(* IEC 61131-3 sources: plc-process-lib/tests/POUs/Suites/FB_Motor_Test, 58 files *)

(* ---- AutoRunStartsAndConfirms.method.decl.st ---- *)
// Auto: запрос xAutoRun запускает двигатель (Starting, xQRun), ОС через 1 с подтверждает пуск (Running);
// пуск считается по фронту ОС, отметка в окне пусков — при входе в Starting; двигатель доступен автоматике.
METHOD PRIVATE AutoRunStartsAndConfirms
VAR
    fbTime   : FB_FakeTime;       // подменное время, старт 1 ч
    fbMot    : FB_Motor;          // двигатель под тестом
    stCmd    : ST_MotorCmd;       // команды
    stRetain : ST_DeviceRetain;   // энергонезависимые данные
    stCfg    : ST_MotorCfg;       // конфигурация (умолчания)
END_VAR

(* ---- CfgChecksSetEachCfgErrBit.method.decl.st ---- *)
// CheckConfig двигателя: каждая проверка 13.9 даёт свой бит wCfgErr; границы допустимы (30 пусков в час,
// tResetPulse = tResetWindow); без ОС времена ОС не проверяются.
METHOD PRIVATE CfgChecksSetEachCfgErrBit
VAR
    fbTime   : FB_FakeTime;       // подменное время, старт 1 ч
    fbMot    : FB_Motor;          // двигатель под тестом
    stCmd    : ST_MotorCmd;       // команды
    stRetain : ST_DeviceRetain;   // энергонезависимые данные
    stCfg    : ST_MotorCfg;       // конфигурация (умолчания)
    uBad     : U_TestEnumInt;     // значение вне перечисления
END_VAR

(* ---- CurrentRunSecondsCountsAndResetsOnStop.method.decl.st ---- *)
// Текущая непрерывная работа: 65 с работы — CurrentRunSeconds = 65 (и stSts.udiRunCurrent_s); останов — 0;
// новый пуск считает с нуля (3 с), наработка всего продолжается (68 с).
// Источник: tools/reference/motor.py, сценарии current_run_*.
METHOD PRIVATE CurrentRunSecondsCountsAndResetsOnStop
VAR
    fbTime   : FB_FakeTime;       // подменное время, старт 1 ч
    fbMot    : FB_Motor;          // двигатель под тестом
    stCmd    : ST_MotorCmd;       // команды
    stRetain : ST_DeviceRetain;   // энергонезависимые данные
    stCfg    : ST_MotorCfg;       // конфигурация (умолчания)
END_VAR

(* ---- ExtFaultInLocalLatches.method.decl.st ---- *)
// Внешняя авария действует и в Local: отказ фиксируется (Fault); после возврата в Manual отказ остаётся,
// пуск — RejectedFault.
METHOD PRIVATE ExtFaultInLocalLatches
VAR
    fbTime   : FB_FakeTime;       // подменное время, старт 1 ч
    fbMot    : FB_Motor;          // двигатель под тестом
    stCmd    : ST_MotorCmd;       // команды
    stRetain : ST_DeviceRetain;   // энергонезависимые данные
    stCfg    : ST_MotorCfg;       // конфигурация (умолчания)
END_VAR

(* ---- ExtFaultTripsAndResetRejectedWhileActive.method.decl.st ---- *)
// Внешняя авария через фильтр tExtFaultFilter = 200 мс: отказ ExtFault, выходы сняты. Reset при действующей
// причине: Accepted и импульс xQReset сразу, к концу окна tResetWindow = 3 с — второй результат RejectedFault,
// отказ остаётся.
METHOD PRIVATE ExtFaultTripsAndResetRejectedWhileActive
VAR
    fbTime   : FB_FakeTime;       // подменное время, старт 1 ч
    fbMot    : FB_Motor;          // двигатель под тестом
    stCmd    : ST_MotorCmd;       // команды
    stRetain : ST_DeviceRetain;   // энергонезависимые данные
    stCfg    : ST_MotorCfg;       // конфигурация (умолчания)
    uiSeqExp : UINT;              // ожидаемый номер команды
END_VAR

(* ---- FailToStopRaisesHighPriorityAlarm.method.decl.st ---- *)
// ОС не пропала после «Стоп»: отказ FailToStop через tFbStop = 5 с; тревога слота 2 — приоритет High
// (механизм не остановить из ПЛК), в сводке ePrioUnack = High, активен только слот 2.
METHOD PRIVATE FailToStopRaisesHighPriorityAlarm
VAR
    fbTime   : FB_FakeTime;       // подменное время, старт 1 ч
    fbMot    : FB_Motor;          // двигатель под тестом
    stCmd    : ST_MotorCmd;       // команды
    stRetain : ST_DeviceRetain;   // энергонезависимые данные
    stCfg    : ST_MotorCfg;       // конфигурация (умолчания)
    itfAlm   : I_Alarm;           // тревога слота
END_VAR

(* ---- FeedbackDropoutWithinFilterNotCountedAsStart.method.decl.st ---- *)
// Дребезг блок-контакта в работе: ОС пропала на 0,2 с (меньше tFbLossFilter = 0,5 с) и вернулась — это не
// останов и не новый пуск: пусков 1, текущая непрерывная работа не обнулилась (по ней станция ограничивает
// непрерывную работу и чередует насосы), отказа нет. Источник: tools/reference/motor.py, сценарии
// dropout_bridged_at_return_s, dropout_bridged_total_s.
METHOD PRIVATE FeedbackDropoutWithinFilterNotCountedAsStart
VAR
    fbTime   : FB_FakeTime;       // подменное время, старт 1 ч
    fbMot    : FB_Motor;          // двигатель под тестом
    stCmd    : ST_MotorCmd;       // команды
    stRetain : ST_DeviceRetain;   // энергонезависимые данные
    stCfg    : ST_MotorCfg;       // конфигурация (умолчания)
END_VAR

(* ---- FeedbackLostWhileRunningTripsAndLatches.method.decl.st ---- *)
// ОС пропала в работе: отказ FeedbackLost через tFbLossFilter = 500 мс (на 400 мс — ещё нет); отказ
// фиксируется — возврат ОС его не снимает, выходы остаются снятыми до Reset.
METHOD PRIVATE FeedbackLostWhileRunningTripsAndLatches
VAR
    fbTime   : FB_FakeTime;       // подменное время, старт 1 ч
    fbMot    : FB_Motor;          // двигатель под тестом
    stCmd    : ST_MotorCmd;       // команды
    stRetain : ST_DeviceRetain;   // энергонезависимые данные
    stCfg    : ST_MotorCfg;       // конфигурация (умолчания)
END_VAR

(* ---- FeedbackStaysAfterTripRaisesFailToStop.method.decl.st ---- *)
// Сварившийся контактор: внешняя авария (тепловое реле) отключила двигатель — xQRun снят, Fault, — а ОС «в
// работе» осталась. Через tFbStop = 5 с после отказа к ExtFault добавляется FailToStop (тревога слота 2, High:
// механизм не остановить из ПЛК); через 4,9 с после отказа — только ExtFault.
METHOD PRIVATE FeedbackStaysAfterTripRaisesFailToStop
VAR
    fbTime   : FB_FakeTime;       // подменное время, старт 1 ч
    fbMot    : FB_Motor;          // двигатель под тестом
    stCmd    : ST_MotorCmd;       // команды
    stRetain : ST_DeviceRetain;   // энергонезависимые данные
    stCfg    : ST_MotorCfg;       // конфигурация (умолчания)
    itfAlm   : I_Alarm;           // тревога слота FailToStop
END_VAR

(* ---- FirstCallSetsTypeSlotsAndPassesDefaultCfg.method.decl.st ---- *)
// Чек-лист устройства, пункты 1 и 4: первый вызов — тип Motor, 8 слотов тревог, умолчания Cfg проходят
// CheckConfig; двигатель стоит, первопричины нет, NE 107 — Good (Manual у двигателя — не CheckFunction).
METHOD PRIVATE FirstCallSetsTypeSlotsAndPassesDefaultCfg
VAR
    fbTime   : FB_FakeTime;       // подменное время, старт 1 ч
    fbMot    : FB_Motor;          // двигатель под тестом
    stCmd    : ST_MotorCmd;       // команды
    stRetain : ST_DeviceRetain;   // энергонезависимые данные
    stCfg    : ST_MotorCfg;       // конфигурация (умолчания)
END_VAR

(* ---- InterlockClearedAutoRestartsManualDoesNot.method.decl.st ---- *)
// Блокировка не фиксируется: в Auto после её снятия двигатель сам запускается по xAutoRun (tMinStop = 0),
// в Manual — нет (ручная защёлка снята блокировкой).
METHOD PRIVATE InterlockClearedAutoRestartsManualDoesNot
VAR
    fbTime    : FB_FakeTime;       // подменное время, старт 1 ч
    fbMot     : FB_Motor;          // двигатель под тестом
    stCmd     : ST_MotorCmd;       // команды
    stRetain  : ST_DeviceRetain;   // энергонезависимые данные
    stCfg     : ST_MotorCfg;       // конфигурация (умолчания)
    fbTime2   : FB_FakeTime;       // подменное время второго двигателя
    fbMot2    : FB_Motor;          // второй двигатель
    stCmd2    : ST_MotorCmd;       // его команды
    stRetain2 : ST_DeviceRetain;   // его энергонезависимые данные
END_VAR

(* ---- InterlockMaskBitClearedIgnored.method.decl.st ---- *)
// Бит блокировки, снятый в wInterlockMask, не действует: двигатель работает, в wInterlock состояния его нет,
// первопричины нет; немаскированный бит останавливает (первопричина — он).
METHOD PRIVATE InterlockMaskBitClearedIgnored
VAR
    fbTime   : FB_FakeTime;       // подменное время, старт 1 ч
    fbMot    : FB_Motor;          // двигатель под тестом
    stCmd    : ST_MotorCmd;       // команды
    stRetain : ST_DeviceRetain;   // энергонезависимые данные
    stCfg    : ST_MotorCfg;       // конфигурация (умолчания)
END_VAR

(* ---- InterlockStopsInAutoAndManualRecordsFirstOut.method.decl.st ---- *)
// Блокировка останавливает двигатель в Auto и в Manual; первопричина — младший из битов, взведённых при
// переходе слова из 0 (биты 3 и 5 разом → 3), последующие биты её не меняют; вход в Starting её снимает;
// в Manual блокировка снимает ручную защёлку.
METHOD PRIVATE InterlockStopsInAutoAndManualRecordsFirstOut
VAR
    fbTime   : FB_FakeTime;       // подменное время, старт 1 ч
    fbMot    : FB_Motor;          // двигатель под тестом
    stCmd    : ST_MotorCmd;       // команды
    stRetain : ST_DeviceRetain;   // энергонезависимые данные
    stCfg    : ST_MotorCfg;       // конфигурация (умолчания)
END_VAR

(* ---- InterlockTripSlotAlarmWhileInterlockActive.method.decl.st ---- *)
// Останов блокировкой в работе — тревога слота 5 InterlockTrip (приоритет по умолчанию None, здесь Low),
// номер тревоги udiAlarmIdBase + 5; пока блокировка действует — тревога активна, после снятия — нет.
METHOD PRIVATE InterlockTripSlotAlarmWhileInterlockActive
VAR
    fbTime   : FB_FakeTime;       // подменное время, старт 1 ч
    fbMot    : FB_Motor;          // двигатель под тестом
    stCmd    : ST_MotorCmd;       // команды
    stRetain : ST_DeviceRetain;   // энергонезависимые данные
    stCfg    : ST_MotorCfg;       // конфигурация (умолчания)
    itfAlm   : I_Alarm;           // тревога слота
END_VAR

(* ---- InvalidCfgAtRuntimeKeepsRunningWithLastValid.method.decl.st ---- *)
// Cfg испорчена в работе (tResetWindow = T#0S): двигатель продолжает работать, CheckFunction и бит
// MOT_CFG_RESET; логика — по последней корректной копии: фильтр пропадания ОС 500 мс, а не 5 с из новой Cfg.
METHOD PRIVATE InvalidCfgAtRuntimeKeepsRunningWithLastValid
VAR
    fbTime   : FB_FakeTime;       // подменное время, старт 1 ч
    fbMot    : FB_Motor;          // двигатель под тестом
    stCmd    : ST_MotorCmd;       // команды
    stRetain : ST_DeviceRetain;   // энергонезависимые данные
    stCfg    : ST_MotorCfg;       // конфигурация (умолчания)
END_VAR

(* ---- InvalidCfgAtStartupStaysStoppedCheckFunction.method.decl.st ---- *)
// Неверная Cfg с первого вызова (uiMaxStartsPerHour > STARTS_WINDOW_MAX): бит MOT_CFG_STARTS_LIMIT,
// CheckFunction, безопасный выход — запрос Auto не запускает, Available = FALSE, xStart — RejectedCfg.
METHOD PRIVATE InvalidCfgAtStartupStaysStoppedCheckFunction
VAR
    fbTime   : FB_FakeTime;       // подменное время, старт 1 ч
    fbMot    : FB_Motor;          // двигатель под тестом
    stCmd    : ST_MotorCmd;       // команды
    stRetain : ST_DeviceRetain;   // энергонезависимые данные
    stCfg    : ST_MotorCfg;       // конфигурация (умолчания)
END_VAR

(* ---- LocalModeOutputsOffTracksFeedback.method.decl.st ---- *)
// Local: выходы сняты, состояние следует ОС (Running/Stopped), контроля ОС нет (ни FailToStop, ни
// UncommandedRun), команды оператора — RejectedMode, блокировка — только предупреждение INTERLOCK_IN_LOCAL.
METHOD PRIVATE LocalModeOutputsOffTracksFeedback
VAR
    fbTime   : FB_FakeTime;       // подменное время, старт 1 ч
    fbMot    : FB_Motor;          // двигатель под тестом
    stCmd    : ST_MotorCmd;       // команды
    stRetain : ST_DeviceRetain;   // энергонезависимые данные
    stCfg    : ST_MotorCfg;       // конфигурация (умолчания)
END_VAR

(* ---- LocalToRemoteRestoresRememberedMode.method.decl.st ---- *)
// Возврат из Local — в запомненный дистанционный режим: Auto → Local → Auto; в Local команда xSetManual меняет
// запомненный режим, и двигатель, запущенный по месту, после возврата продолжает работать в Manual.
METHOD PRIVATE LocalToRemoteRestoresRememberedMode
VAR
    fbTime   : FB_FakeTime;       // подменное время, старт 1 ч
    fbMot    : FB_Motor;          // двигатель под тестом
    stCmd    : ST_MotorCmd;       // команды
    stRetain : ST_DeviceRetain;   // энергонезависимые данные
    stCfg    : ST_MotorCfg;       // конфигурация (умолчания)
END_VAR

(* ---- MaintIntervalReachedMaintenanceRequired.method.decl.st ---- *)
// ТО по наработке 1 ч (порог 3600 с) и по 2 пускам: 3590 с + 10 с работы — предупреждение MAINT_RUNTIME,
// NE 107 MaintenanceRequired; второй пуск — MAINT_STARTS; xResetMaint обнуляет счётчики «с ТО» (Accepted).
// Источник: tools/reference/motor.py, сценарии maint_runtime_*.
METHOD PRIVATE MaintIntervalReachedMaintenanceRequired
VAR
    fbTime   : FB_FakeTime;       // подменное время, старт 1 ч
    fbMot    : FB_Motor;          // двигатель под тестом
    stCmd    : ST_MotorCmd;       // команды
    stRetain : ST_DeviceRetain;   // энергонезависимые данные
    stCfg    : ST_MotorCfg;       // конфигурация (умолчания)
END_VAR

(* ---- ManualStartFeedbackOkGoesRunning.method.decl.st ---- *)
// Manual: xStart принимается (Accepted, импульс сброшен), двигатель в Starting ждёт ОС; ОС через 2 с (меньше
// tFbStart = 5 с) — Running без отказа.
METHOD PRIVATE ManualStartFeedbackOkGoesRunning
VAR
    fbTime   : FB_FakeTime;       // подменное время, старт 1 ч
    fbMot    : FB_Motor;          // двигатель под тестом
    stCmd    : ST_MotorCmd;       // команды
    stRetain : ST_DeviceRetain;   // энергонезависимые данные
    stCfg    : ST_MotorCfg;       // конфигурация (умолчания)
END_VAR

(* ---- ManualStartInAutoRejected.method.decl.st ---- *)
// Auto: команда оператора «Пуск» отклоняется (RejectedMode), импульс сброшен, двигатель стоит, режим Auto.
METHOD PRIVATE ManualStartInAutoRejected
VAR
    fbTime   : FB_FakeTime;       // подменное время, старт 1 ч
    fbMot    : FB_Motor;          // двигатель под тестом
    stCmd    : ST_MotorCmd;       // команды
    stRetain : ST_DeviceRetain;   // энергонезависимые данные
    stCfg    : ST_MotorCfg;       // конфигурация (умолчания)
END_VAR

(* ---- ManualStartRejectionReasonByPrecedence.method.decl.st ---- *)
// Причина отказа xStart в Manual — по старшинству 13.5: при отказе, блокировке, нет разрешения и паузе —
// RejectedFault; без отказа — RejectedInterlock; без блокировки — RejectedPermit; затем RejectedInhibit.
METHOD PRIVATE ManualStartRejectionReasonByPrecedence
VAR
    fbTime   : FB_FakeTime;       // подменное время, старт 1 ч
    fbMot    : FB_Motor;          // двигатель под тестом
    stCmd    : ST_MotorCmd;       // команды
    stRetain : ST_DeviceRetain;   // энергонезависимые данные
    stCfg    : ST_MotorCfg;       // конфигурация (умолчания)
END_VAR

(* ---- MinRunTimeDelaysAutoStop.method.decl.st ---- *)
// tMinRun = 10 с: снятие xAutoRun через 2 с после входа в Running останавливает двигатель только через 10 с
// от входа в Running (на 9,9 с ещё работает).
METHOD PRIVATE MinRunTimeDelaysAutoStop
VAR
    fbTime   : FB_FakeTime;       // подменное время, старт 1 ч
    fbMot    : FB_Motor;          // двигатель под тестом
    stCmd    : ST_MotorCmd;       // команды
    stRetain : ST_DeviceRetain;   // энергонезависимые данные
    stCfg    : ST_MotorCfg;       // конфигурация (умолчания)
END_VAR

(* ---- MinRunTimeManualStopImmediate.method.decl.st ---- *)
// tMinRun действует только на остановы от автоматики: «Стоп» оператора через 1 с после пуска снимает команду
// сразу; в Auto блокировка тоже останавливает без ожидания tMinRun.
METHOD PRIVATE MinRunTimeManualStopImmediate
VAR
    fbTime    : FB_FakeTime;       // подменное время, старт 1 ч
    fbMot     : FB_Motor;          // двигатель под тестом
    stCmd     : ST_MotorCmd;       // команды
    stRetain  : ST_DeviceRetain;   // энергонезависимые данные
    stCfg     : ST_MotorCfg;       // конфигурация (умолчания)
    fbTime2   : FB_FakeTime;       // подменное время второго двигателя
    fbMot2    : FB_Motor;          // второй двигатель
    stCmd2    : ST_MotorCmd;       // его команды
    stRetain2 : ST_DeviceRetain;   // его энергонезависимые данные
END_VAR

(* ---- MinStopTimeInhibitsRestartReportsRemaining.method.decl.st ---- *)
// tMinStop = 30 с: пауза отсчитывается от старта ПЛК и от останова; остаток — в uiInhibitRemain_s с
// округлением вверх (30, через 12,3 с — 18, через 29,9 с — 1), бит START_INHIBIT, xStart — RejectedInhibit;
// через 30 с пуск принимается. Источник: tools/reference/motor.py, сценарии inhibit_min_stop_*.
METHOD PRIVATE MinStopTimeInhibitsRestartReportsRemaining
VAR
    fbTime   : FB_FakeTime;       // подменное время, старт 1 ч
    fbMot    : FB_Motor;          // двигатель под тестом
    stCmd    : ST_MotorCmd;       // команды
    stRetain : ST_DeviceRetain;   // энергонезависимые данные
    stCfg    : ST_MotorCfg;       // конфигурация (умолчания)
END_VAR

(* ---- ModeAutoToManualBumpless.method.decl.st ---- *)
// Auto → Manual при работе: ручная защёлка := команда работы, двигатель продолжает работать; снятие xAutoRun в
// Manual его не останавливает.
METHOD PRIVATE ModeAutoToManualBumpless
VAR
    fbTime   : FB_FakeTime;       // подменное время, старт 1 ч
    fbMot    : FB_Motor;          // двигатель под тестом
    stCmd    : ST_MotorCmd;       // команды
    stRetain : ST_DeviceRetain;   // энергонезависимые данные
    stCfg    : ST_MotorCfg;       // конфигурация (умолчания)
END_VAR

(* ---- NoFeedbackConfiguredRunsOnCommand.method.decl.st ---- *)
// Без ОС (xFbUsed = FALSE; tFbStart = T#0S тогда допустим): работа — по команде, сразу Running; отказов
// контроля ОС нет; наработка и пуски — по команде.
METHOD PRIVATE NoFeedbackConfiguredRunsOnCommand
VAR
    fbTime   : FB_FakeTime;       // подменное время, старт 1 ч
    fbMot    : FB_Motor;          // двигатель под тестом
    stCmd    : ST_MotorCmd;       // команды
    stRetain : ST_DeviceRetain;   // энергонезависимые данные
    stCfg    : ST_MotorCfg;       // конфигурация (умолчания)
END_VAR

(* ---- NoFeedbackSetsFailToStartAfterTimeout.method.decl.st ---- *)
// Нет ОС после пуска: отказ FailToStart ровно через tFbStart = 5 с (на 4,9 с — ещё нет), выходы сняты, Fault,
// NE 107 Failure, тревога слота 0 активна и не квитирована.
METHOD PRIVATE NoFeedbackSetsFailToStartAfterTimeout
VAR
    fbTime   : FB_FakeTime;       // подменное время, старт 1 ч
    fbMot    : FB_Motor;          // двигатель под тестом
    stCmd    : ST_MotorCmd;       // команды
    stRetain : ST_DeviceRetain;   // энергонезависимые данные
    stCfg    : ST_MotorCfg;       // конфигурация (умолчания)
    itfAlm   : I_Alarm;           // тревога слота
END_VAR

(* ---- OosEntryClearsLatchedFaultsAndFirstOut.method.decl.st ---- *)
// Чек-лист, пункт 5: вход в OutOfService (хук OnModeChanged) снимает зафиксированный отказ и первопричину;
// тревоги — OutOfService, NE 107 — CheckFunction.
METHOD PRIVATE OosEntryClearsLatchedFaultsAndFirstOut
VAR
    fbTime   : FB_FakeTime;       // подменное время, старт 1 ч
    fbMot    : FB_Motor;          // двигатель под тестом
    stCmd    : ST_MotorCmd;       // команды
    stRetain : ST_DeviceRetain;   // энергонезависимые данные
    stCfg    : ST_MotorCfg;       // конфигурация (умолчания)
    itfAlm   : I_Alarm;           // тревога слота
END_VAR

(* ---- OosRequestWhileRunningByFeedbackRejected.method.decl.st ---- *)
// Вывод из работы — только когда механизм стоит (2.2): после внешней аварии команда снята (Fault), но ОС
// «в работе» держится (сварился контактор) — xSetOos отклоняется (RejectedState), зафиксированные отказы не
// снимаются; ОС пропала — вывод из работы принят.
METHOD PRIVATE OosRequestWhileRunningByFeedbackRejected
VAR
    fbTime   : FB_FakeTime;       // подменное время, старт 1 ч
    fbMot    : FB_Motor;          // двигатель под тестом
    stCmd    : ST_MotorCmd;       // команды
    stRetain : ST_DeviceRetain;   // энергонезависимые данные
    stCfg    : ST_MotorCfg;       // конфигурация (умолчания)
END_VAR

(* ---- OosRequestWhileRunningRejected.method.decl.st ---- *)
// Вывод из работы при работающем двигателе — RejectedState (чек-лист, пункт 3); у стоящего — принят: режим
// OutOfService, NE 107 CheckFunction, пуск — RejectedMode.
METHOD PRIVATE OosRequestWhileRunningRejected
VAR
    fbTime   : FB_FakeTime;       // подменное время, старт 1 ч
    fbMot    : FB_Motor;          // двигатель под тестом
    stCmd    : ST_MotorCmd;       // команды
    stRetain : ST_DeviceRetain;   // энергонезависимые данные
    stCfg    : ST_MotorCfg;       // конфигурация (умолчания)
END_VAR

(* ---- PermitMissingBlocksStartDoesNotStopRunning.method.decl.st ---- *)
// Нет разрешения: в Auto запрос ждёт (бит PERMIT_MISSING, wPermitMissing, ReadyToStart = FALSE) и пуск
// происходит сам, когда разрешение появилось; пропажа разрешения работающий двигатель не останавливает;
// в Manual xStart — RejectedPermit.
METHOD PRIVATE PermitMissingBlocksStartDoesNotStopRunning
VAR
    fbTime    : FB_FakeTime;       // подменное время, старт 1 ч
    fbMot     : FB_Motor;          // двигатель под тестом
    stCmd     : ST_MotorCmd;       // команды
    stRetain  : ST_DeviceRetain;   // энергонезависимые данные
    stCfg     : ST_MotorCfg;       // конфигурация (умолчания)
    fbTime2   : FB_FakeTime;       // подменное время второго двигателя
    fbMot2    : FB_Motor;          // второй двигатель
    stCmd2    : ST_MotorCmd;       // его команды
    stRetain2 : ST_DeviceRetain;   // его энергонезависимые данные
END_VAR

(* ---- PlcRestartAutoWithoutDemandStops.method.decl.st ---- *)
// Старт ПЛК в Auto без запроса при работающем по ОС двигателе: штатный останов с контролем (Stopping, команда
// не подаётся), после пропадания ОС — Stopped без отказа.
METHOD PRIVATE PlcRestartAutoWithoutDemandStops
VAR
    fbTime   : FB_FakeTime;       // подменное время, старт 1 ч
    fbMot    : FB_Motor;          // двигатель под тестом
    stCmd    : ST_MotorCmd;       // команды
    stRetain : ST_DeviceRetain;   // энергонезависимые данные
    stCfg    : ST_MotorCfg;       // конфигурация (умолчания)
END_VAR

(* ---- PlcRestartRunningFeedbackAdopted.method.decl.st ---- *)
// Старт ПЛК при работающем по ОС двигателе: Auto с запросом и Manual — подхват (Running, xQRun) без отказа
// UncommandedRun и без счёта пуска.
METHOD PRIVATE PlcRestartRunningFeedbackAdopted
VAR
    fbTime    : FB_FakeTime;       // подменное время, старт 1 ч
    fbMot     : FB_Motor;          // двигатель под тестом
    stCmd     : ST_MotorCmd;       // команды
    stRetain  : ST_DeviceRetain;   // энергонезависимые данные
    stCfg     : ST_MotorCfg;       // конфигурация (умолчания)
    fbTime2   : FB_FakeTime;       // подменное время второго двигателя
    fbMot2    : FB_Motor;          // второй двигатель
    stCmd2    : ST_MotorCmd;       // его команды
    stRetain2 : ST_DeviceRetain;   // его энергонезависимые данные
END_VAR

(* ---- PowerDipFeedbackStaysStoppingWithoutUncommandedRun.method.decl.st ---- *)
// Провал напряжения 0,3 с, который пережил ПЧ (кинетическая поддержка): ОС «в работе» не пропала. Команда
// снята; после восстановления питания двигатель тормозит под контролем останова (Stopping, tFbStop = 10 с), а
// не стоит в Stopped с ложным UncommandedRun через tFbStart = 5 с; ОС пропала через 6 с — Stopped без отказа.
METHOD PRIVATE PowerDipFeedbackStaysStoppingWithoutUncommandedRun
VAR
    fbTime   : FB_FakeTime;       // подменное время, старт 1 ч
    fbMot    : FB_Motor;          // двигатель под тестом
    stCmd    : ST_MotorCmd;       // команды
    stRetain : ST_DeviceRetain;   // энергонезависимые данные
    stCfg    : ST_MotorCfg;       // конфигурация
END_VAR

(* ---- PowerDipWhileStoppedPauseFromPowerLoss.method.decl.st ---- *)
// Провал питания у стоящего двигателя тоже даёт паузу tMinStop = 20 с от момента пропадания: через 5 с после
// провала (питание вернулось через 1 с) пуск — RejectedInhibit, остаток 15 с; через 20 с — принят.
// Источник: tools/reference/motor.py, сценарий inhibit_power_loss_after_5s.
METHOD PRIVATE PowerDipWhileStoppedPauseFromPowerLoss
VAR
    fbTime   : FB_FakeTime;       // подменное время, старт 1 ч
    fbMot    : FB_Motor;          // двигатель под тестом
    stCmd    : ST_MotorCmd;       // команды
    stRetain : ST_DeviceRetain;   // энергонезависимые данные
    stCfg    : ST_MotorCfg;       // конфигурация (умолчания)
END_VAR

(* ---- PowerLossInManualLatchClearedNoRestart.method.decl.st ---- *)
// Пропадание напряжения в Manual снимает ручную защёлку: после восстановления питания двигатель не
// запускается сам; отказа нет.
METHOD PRIVATE PowerLossInManualLatchClearedNoRestart
VAR
    fbTime   : FB_FakeTime;       // подменное время, старт 1 ч
    fbMot    : FB_Motor;          // двигатель под тестом
    stCmd    : ST_MotorCmd;       // команды
    stRetain : ST_DeviceRetain;   // энергонезависимые данные
    stCfg    : ST_MotorCfg;       // конфигурация (умолчания)
END_VAR

(* ---- PowerLossStopsWithoutFaultStartsMinStop.method.decl.st ---- *)
// Пропадание напряжения в Auto: Stopped без отказа, предупреждение POWER_LOST и запрет пуска; tMinStop = 20 с
// отсчитывается от момента пропадания: питание вернулось через 5 с — остаток 15 с, пуск по запросу Auto — ровно
// через 20 с. Источник: tools/reference/motor.py, сценарий inhibit_power_loss_after_5s.
METHOD PRIVATE PowerLossStopsWithoutFaultStartsMinStop
VAR
    fbTime   : FB_FakeTime;       // подменное время, старт 1 ч
    fbMot    : FB_Motor;          // двигатель под тестом
    stCmd    : ST_MotorCmd;       // команды
    stRetain : ST_DeviceRetain;   // энергонезависимые данные
    stCfg    : ST_MotorCfg;       // конфигурация (умолчания)
END_VAR

(* ---- PresetCountersAppliedInBody.method.decl.st ---- *)
// PresetCounters() только ставит запрос (TRUE), значения пишет ближайший вызов тела: наработка и пуски в
// stRetain, RunSeconds, Starts, rRunTime_h = 100 ч, Accepted; счётчики «с ТО» не меняются.
METHOD PRIVATE PresetCountersAppliedInBody
VAR
    fbTime   : FB_FakeTime;       // подменное время, старт 1 ч
    fbMot    : FB_Motor;          // двигатель под тестом
    stCmd    : ST_MotorCmd;       // команды
    stRetain : ST_DeviceRetain;   // энергонезависимые данные
    stCfg    : ST_MotorCfg;       // конфигурация (умолчания)
END_VAR

(* ---- ReadyToStartFalseWhileStarting.method.decl.st ---- *)
// ReadyToStart — «стоит и готов к пуску» (I_Motor): в Auto до пуска TRUE; в Starting (команда подана, ОС ещё
// нет, tMinStop = 0) — FALSE: станция не должна считать запускаемый насос резервом; в Running — FALSE.
METHOD PRIVATE ReadyToStartFalseWhileStarting
VAR
    fbTime   : FB_FakeTime;       // подменное время, старт 1 ч
    fbMot    : FB_Motor;          // двигатель под тестом
    stCmd    : ST_MotorCmd;       // команды
    stRetain : ST_DeviceRetain;   // энергонезависимые данные
    stCfg    : ST_MotorCfg;       // конфигурация (умолчания)
END_VAR

(* ---- ResetCauseClearsWithinWindowFaultCleared.method.decl.st ---- *)
// Reset при действующей причине, причина уходит через 1 с (в окне tResetWindow = 3 с): отказ снимается без
// второго нажатия, двигатель Stopped; RejectedFault в конце окна не появляется.
METHOD PRIVATE ResetCauseClearsWithinWindowFaultCleared
VAR
    fbTime   : FB_FakeTime;       // подменное время, старт 1 ч
    fbMot    : FB_Motor;          // двигатель под тестом
    stCmd    : ST_MotorCmd;       // команды
    stRetain : ST_DeviceRetain;   // энергонезависимые данные
    stCfg    : ST_MotorCfg;       // конфигурация (умолчания)
    uiSeqExp : UINT;              // номер команды после Reset
END_VAR

(* ---- ResetFailToStopClearedOnlyAfterMotorStops.method.decl.st ---- *)
// FailToStop снимается Reset только когда двигатель не работает по ОС (M-02): Reset при ещё работающем
// двигателе — импульс xQReset, отказ остаётся, к концу окна tResetWindow = 3 с второй результат RejectedFault;
// ОС пропала — следующий Reset снимает отказ, двигатель в Stopped.
METHOD PRIVATE ResetFailToStopClearedOnlyAfterMotorStops
VAR
    fbTime   : FB_FakeTime;       // подменное время, старт 1 ч
    fbMot    : FB_Motor;          // двигатель под тестом
    stCmd    : ST_MotorCmd;       // команды
    stRetain : ST_DeviceRetain;   // энергонезависимые данные
    stCfg    : ST_MotorCfg;       // конфигурация (умолчания)
END_VAR

(* ---- ResetPulsesResetOutput.method.decl.st ---- *)
// Reset без отказов (чек-лист, пункт 2): результат Accepted, uiCmdSeq + 1; импульс xQReset длится
// tResetPulse = 1 с (на 0,9 с ещё есть, на 1,0 с — нет); RejectedFault в конце окна нет.
METHOD PRIVATE ResetPulsesResetOutput
VAR
    fbTime   : FB_FakeTime;       // подменное время, старт 1 ч
    fbMot    : FB_Motor;          // двигатель под тестом
    stCmd    : ST_MotorCmd;       // команды
    stRetain : ST_DeviceRetain;   // энергонезависимые данные
    stCfg    : ST_MotorCfg;       // конфигурация (умолчания)
    uiSeqExp : UINT;              // ожидаемый номер команды
END_VAR

(* ---- RunHoursAccumulateInRetain.method.decl.st ---- *)
// Наработка копится в stRetain: 90 мин работы шагами по 10 с — 5400 с, rRunTime_h = 1,5 ч (и «с ТО» так же,
// RunSeconds); 2,5 с шагами по 100 мс — 2 целых секунды (0,5 с — в накопителе), ещё 0,5 с — 3 с.
// Источник: tools/reference/motor.py, сценарии run_hours_90min_*, run_fraction_*.
METHOD PRIVATE RunHoursAccumulateInRetain
VAR
    fbTime    : FB_FakeTime;       // подменное время, старт 1 ч
    fbMot     : FB_Motor;          // двигатель под тестом
    stCmd     : ST_MotorCmd;       // команды
    stRetain  : ST_DeviceRetain;   // энергонезависимые данные
    stCfg     : ST_MotorCfg;       // конфигурация (умолчания)
    fbTime2   : FB_FakeTime;       // подменное время второго двигателя
    fbMot2    : FB_Motor;          // второй двигатель
    stCmd2    : ST_MotorCmd;       // его команды
    stRetain2 : ST_DeviceRetain;   // его энергонезависимые данные
END_VAR

(* ---- RunHoursLargeTimeStepBounded.method.decl.st ---- *)
// Шаг времени больше DT_ACCUM_MAX (зависание, остановка задачи) засчитывается как 10 с: после шага 1 ч — 10 с,
// после шага 3 с — 13 с. Источник: tools/reference/motor.py, сценарии run_large_step_*.
METHOD PRIVATE RunHoursLargeTimeStepBounded
VAR
    fbTime   : FB_FakeTime;       // подменное время, старт 1 ч
    fbMot    : FB_Motor;          // двигатель под тестом
    stCmd    : ST_MotorCmd;       // команды
    stRetain : ST_DeviceRetain;   // энергонезависимые данные
    stCfg    : ST_MotorCfg;       // конфигурация (умолчания)
END_VAR

(* ---- SetSlotPriority.method.decl.st ---- *)
// Помощник: приоритет слота тревоги в Cfg двигателя (через копию элемента)
METHOD PRIVATE SetSlotPriority
VAR_IN_OUT
    stCfgMot : ST_MotorCfg;         // конфигурация двигателя
END_VAR
VAR_INPUT
    uiSlot    : UINT;               // номер слота
    ePrioSlot : E_AlarmPriority;    // приоритет
END_VAR
VAR
    stSlot : ST_AlarmCfg;           // копия слота
END_VAR

(* ---- Spin.method.decl.st ---- *)
// Помощник: uiN вызовов двигателя, перед каждым — шаг подменного времени tDt (T#0S — тот же момент).
// Входы двигателя тест пишет по имени экземпляра до вызова помощника; ассертов внутри нет
METHOD PRIVATE Spin
VAR_IN_OUT
    fbM : FB_Motor;          // двигатель
    fbT : FB_FakeTime;       // подменное время
    stC : ST_MotorCmd;       // команды
    stR : ST_DeviceRetain;   // энергонезависимые данные
END_VAR
VAR_IN_OUT CONSTANT
    stF : ST_MotorCfg;       // конфигурация
END_VAR
VAR_INPUT
    uiN : UINT;              // число вызовов
    tDt : TIME;              // шаг времени перед каждым вызовом
END_VAR
VAR
    uiLoop : UINT;           // номер вызова
END_VAR

(* ---- Spin.method.impl.st ---- *)
FOR uiLoop := 1 TO uiN DO
    fbT.Advance(tStep := tDt);
    fbM(itfTime := fbT, stCmd := stC, stRetain := stR, stCfg := stF);
END_FOR

(* ---- StartsCountedOnFeedbackEdge.method.decl.st ---- *)
// Пуск считается по фронту ОС: попытка пуска без ОС — отметка в окне, но не пуск; ОС — пуск (всего и «с ТО»);
// пуск по месту (фронт ОС в Local без команды ПЛК) — тоже пуск и отметка в окне.
METHOD PRIVATE StartsCountedOnFeedbackEdge
VAR
    fbTime   : FB_FakeTime;       // подменное время, старт 1 ч
    fbMot    : FB_Motor;          // двигатель под тестом
    stCmd    : ST_MotorCmd;       // команды
    stRetain : ST_DeviceRetain;   // энергонезависимые данные
    stCfg    : ST_MotorCfg;       // конфигурация (умолчания)
END_VAR

(* ---- StartsPerHourLimitReachedInhibitsUntilWindowFrees.method.decl.st ---- *)
// Лимит 3 пуска в час, пуски в t0, t0 + 10 мин, t0 + 20 мин: в t0 + 30 мин пуск отклонён (RejectedInhibit),
// uiStartsLastHour = 3, остаток 1800 с, предупреждение STARTS_LIMIT; в t0 + 59 мин остаток 60 с; в t0 + 60 мин
// первая отметка вышла из окна — пуск принят. Источник: tools/reference/motor.py, сценарии starts_limit_3_*.
METHOD PRIVATE StartsPerHourLimitReachedInhibitsUntilWindowFrees
VAR
    fbTime   : FB_FakeTime;       // подменное время, старт 1 ч
    fbMot    : FB_Motor;          // двигатель под тестом
    stCmd    : ST_MotorCmd;       // команды
    stRetain : ST_DeviceRetain;   // энергонезависимые данные
    stCfg    : ST_MotorCfg;       // конфигурация (умолчания)
END_VAR

(* ---- StartWhileStoppingPermitLostCancelsLatch.method.decl.st ---- *)
// Manual: «Пуск» во время выбега (Stopping) принят — двигатель запустится после останова (M-09). За время
// выбега пропало разрешение: после останова отложенный пуск отменяется (защёлка снята, второй результат
// RejectedPermit), и когда разрешение вернётся через 10 мин, двигатель в Manual сам не запускается.
METHOD PRIVATE StartWhileStoppingPermitLostCancelsLatch
VAR
    fbTime   : FB_FakeTime;       // подменное время, старт 1 ч
    fbMot    : FB_Motor;          // двигатель под тестом
    stCmd    : ST_MotorCmd;       // команды
    stRetain : ST_DeviceRetain;   // энергонезависимые данные
    stCfg    : ST_MotorCfg;       // конфигурация (умолчания)
END_VAR

(* ---- StopAndStartSameCallStopWins.method.decl.st ---- *)
// «Стоп» и «Пуск» в одном вызове: «Стоп» старше — двигатель останавливается, оба импульса сброшены.
METHOD PRIVATE StopAndStartSameCallStopWins
VAR
    fbTime   : FB_FakeTime;       // подменное время, старт 1 ч
    fbMot    : FB_Motor;          // двигатель под тестом
    stCmd    : ST_MotorCmd;       // команды
    stRetain : ST_DeviceRetain;   // энергонезависимые данные
    stCfg    : ST_MotorCfg;       // конфигурация (умолчания)
END_VAR

(* ---- StopInAutoSwitchesToManualAndStops.method.decl.st ---- *)
// «Стоп» оператора в Auto: устройство переходит в Manual (запомнено в retain), команда работы снимается сразу,
// Stopping до пропадания ОС, затем Stopped; результат Accepted.
METHOD PRIVATE StopInAutoSwitchesToManualAndStops
VAR
    fbTime   : FB_FakeTime;       // подменное время, старт 1 ч
    fbMot    : FB_Motor;          // двигатель под тестом
    stCmd    : ST_MotorCmd;       // команды
    stRetain : ST_DeviceRetain;   // энергонезависимые данные
    stCfg    : ST_MotorCfg;       // конфигурация (умолчания)
END_VAR

(* ---- TimeBackwardsDuringMinRunKeepsRunning.method.decl.st ---- *)
// Auto, tMinRun = 10 с: через 2 с работы запрос снят — двигатель работает до tMinRun. Время назад на 30 с: отсчёт
// tMinRun начинается заново (M-17), двигатель не останавливается раньше срока; останов ровно через 10 с после скачка.
METHOD PRIVATE TimeBackwardsDuringMinRunKeepsRunning
VAR
    fbTime   : FB_FakeTime;       // подменное время, старт 1 ч
    fbMot    : FB_Motor;          // двигатель под тестом
    stCmd    : ST_MotorCmd;       // команды
    stRetain : ST_DeviceRetain;   // энергонезависимые данные
    stCfg    : ST_MotorCfg;       // конфигурация
END_VAR

(* ---- TimeBackwardsDuringMinStopPauseRestarts.method.decl.st ---- *)
// Пауза tMinStop = 10 с (защита погружного насоса от обратного вращения): двигатель остановлен, прошло 2 с, время
// назад на 30 с (SetNow — смена источника времени). Пауза отсчитывается заново (M-03, M-17), а не снимается
// переполнением LTIME без знака: пуск — RejectedInhibit, остаток 10 с; 1 с в 9,9 с; через 10 с пуск принят.
METHOD PRIVATE TimeBackwardsDuringMinStopPauseRestarts
VAR
    fbTime   : FB_FakeTime;       // подменное время, старт 1 ч
    fbMot    : FB_Motor;          // двигатель под тестом
    stCmd    : ST_MotorCmd;       // команды
    stRetain : ST_DeviceRetain;   // энергонезависимые данные
    stCfg    : ST_MotorCfg;       // конфигурация
END_VAR

(* ---- TimeBackwardsDuringResetPulsePulseRestarts.method.decl.st ---- *)
// Внешняя авария зафиксирована, Reset с tResetPulse = 1 с (сброс УПП): через 0,5 с время назад на 30 с. Импульс
// xQReset и окно tResetWindow отсчитываются заново (M-17), а не обрываются переполнением: импульс держится ещё 1 с
// после скачка; авария, снятая в окне, сброшена без RejectedFault.
METHOD PRIVATE TimeBackwardsDuringResetPulsePulseRestarts
VAR
    fbTime   : FB_FakeTime;       // подменное время, старт 1 ч
    fbMot    : FB_Motor;          // двигатель под тестом
    stCmd    : ST_MotorCmd;       // команды
    stRetain : ST_DeviceRetain;   // энергонезависимые данные
    stCfg    : ST_MotorCfg;       // конфигурация
END_VAR

(* ---- TimeBackwardsNoFaultNoCountJump.method.decl.st ---- *)
// «Время назад» (SetNow на 30 с раньше) у работающего двигателя: отказов нет, наработка не скачет (шаг
// времени 0), дальше считается обычно.
METHOD PRIVATE TimeBackwardsNoFaultNoCountJump
VAR
    fbTime   : FB_FakeTime;       // подменное время, старт 1 ч
    fbMot    : FB_Motor;          // двигатель под тестом
    stCmd    : ST_MotorCmd;       // команды
    stRetain : ST_DeviceRetain;   // энергонезависимые данные
    stCfg    : ST_MotorCfg;       // конфигурация (умолчания)
END_VAR

(* ---- UncommandedRunDetected.method.decl.st ---- *)
// ОС без команды ПЛК дольше tFbStart = 5 с: отказ UncommandedRun (High); до этого двигатель считается
// работающим по ОС; фронт ОС без команды — пуск (счётчик и окно пусков).
METHOD PRIVATE UncommandedRunDetected
VAR
    fbTime   : FB_FakeTime;       // подменное время, старт 1 ч
    fbMot    : FB_Motor;          // двигатель под тестом
    stCmd    : ST_MotorCmd;       // команды
    stRetain : ST_DeviceRetain;   // энергонезависимые данные
    stCfg    : ST_MotorCfg;       // конфигурация (умолчания)
END_VAR
